// SIMATIC S7-200 SMART project (STEP 7-Micro/WIN SMART), CPU ST30

SYMBOL_TABLE System Symbols
Always_On        SM0.0    // Always ON
First_Scan_On    SM0.1    // ON for the first scan cycle only
END_SYMBOL_TABLE

ORGANIZATION_BLOCK MAIN:OB1
TITLE=Program Comments
BEGIN
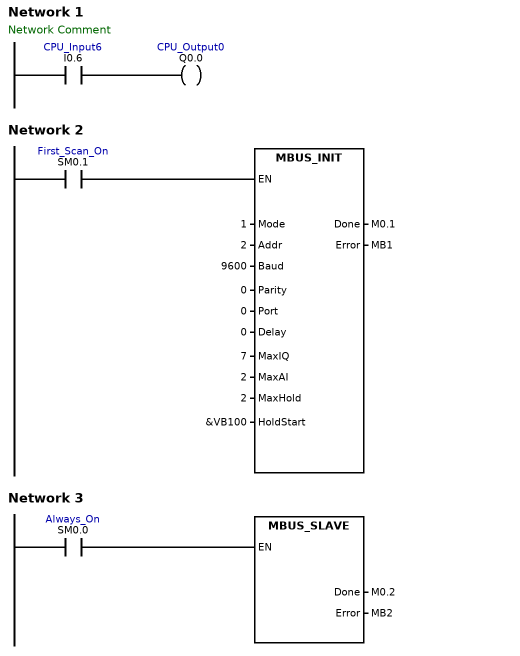
Network 1
// Network Comment
LD     CPU_Input6:I0.6
=      CPU_Output0:Q0.0
Network 2
LD     First_Scan_On:SM0.1
CALL   MBUS_INIT:SBR1, 1, 2, 9600, 0, 0, 0, 7, 2, 2, &VB100, M0.1, MB1
Network 3
LD     Always_On:SM0.0
CALL   MBUS_SLAVE:SBR2, M0.2, MB2
END_ORGANIZATION_BLOCK

// SBR1: protected block, not included

// SBR2: protected block, not included

// SBR3: protected block, not included
